Fanuc KAREL source: kb00168.KL

PROGRAM KB00168
%NOLOCKGROUP
VAR
P1 : STRING[80];P2:INTEGER
BEGIN
--
P1='A'
P2=1
SET_LANG(P1,P2)
END KB00168
